// TIA Portal V18 export
DATA_BLOCK "DB_App"   // DB2
// stored: InstanceOfName FB_App, InstanceOfType FB
"FB_App"
   // VAR
   //    frequencySource_Last : Int;
   //    frequencySetpoint_Last : Real;
   //    state_start : Bool;
   //    state_rev : Bool;
   //    state_stop : Bool;
   //    i : Int;
   //    state_alarm : Bool;
   // END_VAR
BEGIN
END_DATA_BLOCK
